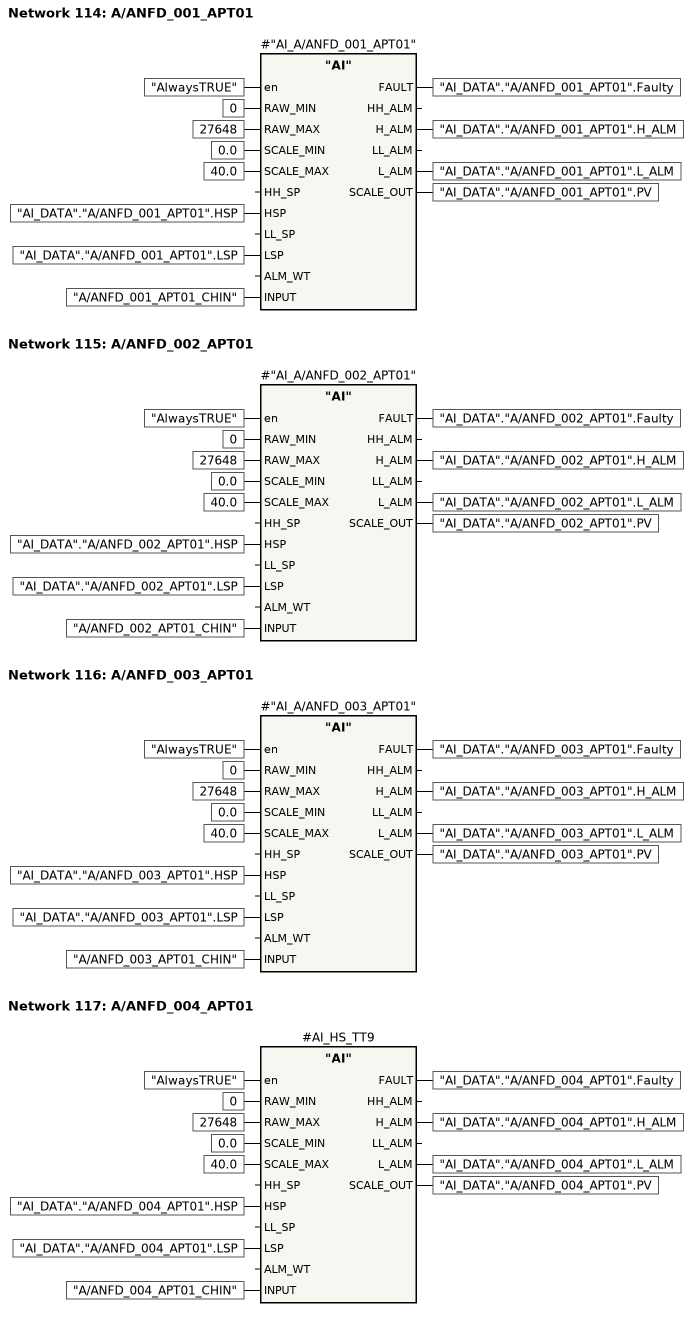
   IF "AlwaysTRUE" THEN
       #"AI_A/ANFD_001_APT01"(RAW_MIN := 0,   // "AI"
                              RAW_MAX := 27648,
                              SCALE_MIN := 0.0,
                              SCALE_MAX := 40.0,
                              HSP := "AI_DATA"."A/ANFD_001_APT01".HSP,
                              LSP := "AI_DATA"."A/ANFD_001_APT01".LSP,
                              INPUT := "A/ANFD_001_APT01_CHIN",
                              FAULT => "AI_DATA"."A/ANFD_001_APT01".Faulty,
                              H_ALM => "AI_DATA"."A/ANFD_001_APT01".H_ALM,
                              L_ALM => "AI_DATA"."A/ANFD_001_APT01".L_ALM,
                              SCALE_OUT => "AI_DATA"."A/ANFD_001_APT01".PV);
   END_IF;
END_REGION

REGION Network 115: A/ANFD_002_APT01
   IF "AlwaysTRUE" THEN
       #"AI_A/ANFD_002_APT01"(RAW_MIN := 0,   // "AI"
                              RAW_MAX := 27648,
                              SCALE_MIN := 0.0,
                              SCALE_MAX := 40.0,
                              HSP := "AI_DATA"."A/ANFD_002_APT01".HSP,
                              LSP := "AI_DATA"."A/ANFD_002_APT01".LSP,
                              INPUT := "A/ANFD_002_APT01_CHIN",
                              FAULT => "AI_DATA"."A/ANFD_002_APT01".Faulty,
                              H_ALM => "AI_DATA"."A/ANFD_002_APT01".H_ALM,
                              L_ALM => "AI_DATA"."A/ANFD_002_APT01".L_ALM,
                              SCALE_OUT => "AI_DATA"."A/ANFD_002_APT01".PV);
   END_IF;
END_REGION

REGION Network 116: A/ANFD_003_APT01
   IF "AlwaysTRUE" THEN
       #"AI_A/ANFD_003_APT01"(RAW_MIN := 0,   // "AI"
                              RAW_MAX := 27648,
                              SCALE_MIN := 0.0,
                              SCALE_MAX := 40.0,
                              HSP := "AI_DATA"."A/ANFD_003_APT01".HSP,
                              LSP := "AI_DATA"."A/ANFD_003_APT01".LSP,
                              INPUT := "A/ANFD_003_APT01_CHIN",
                              FAULT => "AI_DATA"."A/ANFD_003_APT01".Faulty,
                              H_ALM => "AI_DATA"."A/ANFD_003_APT01".H_ALM,
                              L_ALM => "AI_DATA"."A/ANFD_003_APT01".L_ALM,
                              SCALE_OUT => "AI_DATA"."A/ANFD_003_APT01".PV);
   END_IF;
END_REGION

REGION Network 117: A/ANFD_004_APT01
   IF "AlwaysTRUE" THEN
       #AI_HS_TT9(RAW_MIN := 0,   // "AI"
                  RAW_MAX := 27648,
                  SCALE_MIN := 0.0,
                  SCALE_MAX := 40.0,
                  HSP := "AI_DATA"."A/ANFD_004_APT01".HSP,
                  LSP := "AI_DATA"."A/ANFD_004_APT01".LSP,
                  INPUT := "A/ANFD_004_APT01_CHIN",
                  FAULT => "AI_DATA"."A/ANFD_004_APT01".Faulty,
                  H_ALM => "AI_DATA"."A/ANFD_004_APT01".H_ALM,
                  L_ALM => "AI_DATA"."A/ANFD_004_APT01".L_ALM,
                  SCALE_OUT => "AI_DATA"."A/ANFD_004_APT01".PV);
   END_IF;
END_REGION

REGION Network 118: A/ANFD_001_TT01
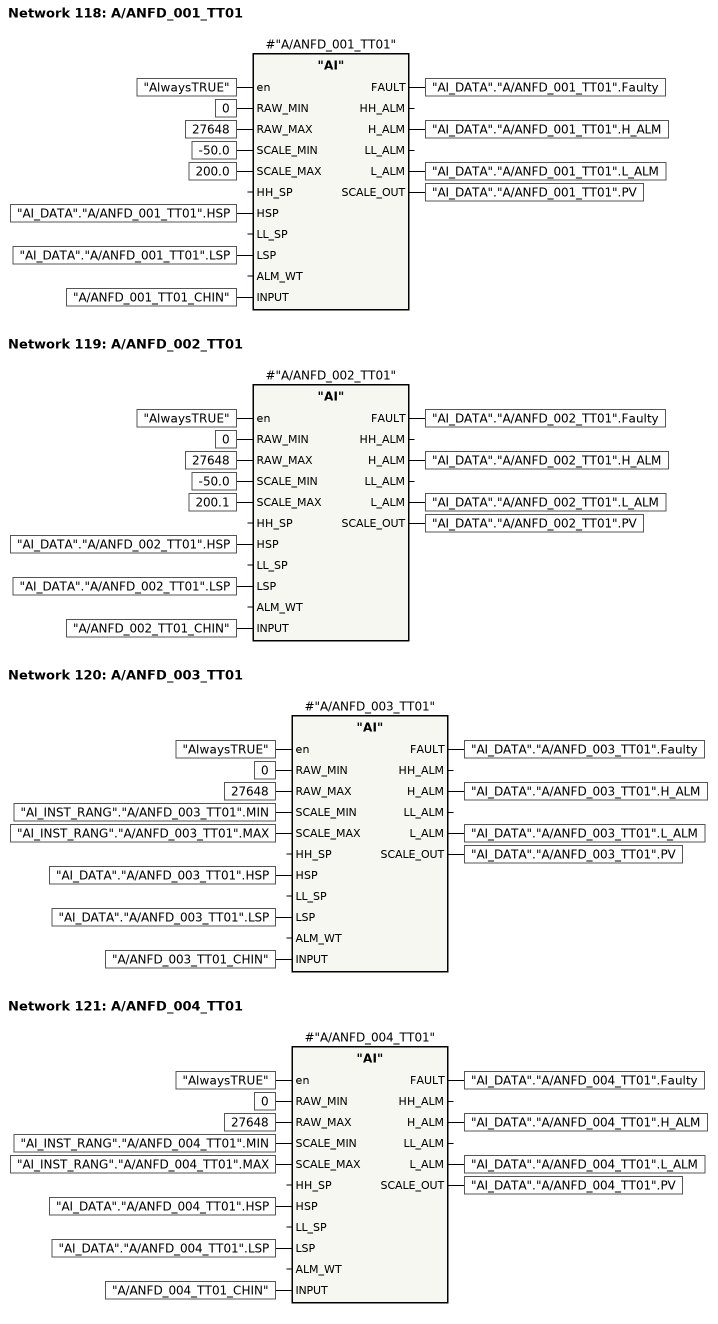
   IF "AlwaysTRUE" THEN
       #"A/ANFD_001_TT01"(RAW_MIN := 0,   // "AI"
                          RAW_MAX := 27648,
                          SCALE_MIN := -50.0,
                          SCALE_MAX := 200.0,
                          HSP := "AI_DATA"."A/ANFD_001_TT01".HSP,
                          LSP := "AI_DATA"."A/ANFD_001_TT01".LSP,
                          INPUT := "A/ANFD_001_TT01_CHIN",
                          FAULT => "AI_DATA"."A/ANFD_001_TT01".Faulty,
                          H_ALM => "AI_DATA"."A/ANFD_001_TT01".H_ALM,
                          L_ALM => "AI_DATA"."A/ANFD_001_TT01".L_ALM,
                          SCALE_OUT => "AI_DATA"."A/ANFD_001_TT01".PV);
   END_IF;
END_REGION

REGION Network 119: A/ANFD_002_TT01
   IF "AlwaysTRUE" THEN
       #"A/ANFD_002_TT01"(RAW_MIN := 0,   // "AI"
                          RAW_MAX := 27648,
                          SCALE_MIN := -50.0,
                          SCALE_MAX := 200.1,
                          HSP := "AI_DATA"."A/ANFD_002_TT01".HSP,
                          LSP := "AI_DATA"."A/ANFD_002_TT01".LSP,
                          INPUT := "A/ANFD_002_TT01_CHIN",
                          FAULT => "AI_DATA"."A/ANFD_002_TT01".Faulty,
                          H_ALM => "AI_DATA"."A/ANFD_002_TT01".H_ALM,
                          L_ALM => "AI_DATA"."A/ANFD_002_TT01".L_ALM,
                          SCALE_OUT => "AI_DATA"."A/ANFD_002_TT01".PV);
   END_IF;
END_REGION

REGION Network 120: A/ANFD_003_TT01
   IF "AlwaysTRUE" THEN
       #"A/ANFD_003_TT01"(RAW_MIN := 0,   // "AI"
                          RAW_MAX := 27648,
                          SCALE_MIN := "AI_INST_RANG"."A/ANFD_003_TT01".MIN,
                          SCALE_MAX := "AI_INST_RANG"."A/ANFD_003_TT01".MAX,
                          HSP := "AI_DATA"."A/ANFD_003_TT01".HSP,
                          LSP := "AI_DATA"."A/ANFD_003_TT01".LSP,
                          INPUT := "A/ANFD_003_TT01_CHIN",
                          FAULT => "AI_DATA"."A/ANFD_003_TT01".Faulty,
                          H_ALM => "AI_DATA"."A/ANFD_003_TT01".H_ALM,
                          L_ALM => "AI_DATA"."A/ANFD_003_TT01".L_ALM,
                          SCALE_OUT => "AI_DATA"."A/ANFD_003_TT01".PV);
   END_IF;
END_REGION

REGION Network 121: A/ANFD_004_TT01
   IF "AlwaysTRUE" THEN
       #"A/ANFD_004_TT01"(RAW_MIN := 0,   // "AI"
                          RAW_MAX := 27648,
                          SCALE_MIN := "AI_INST_RANG"."A/ANFD_004_TT01".MIN,
                          SCALE_MAX := "AI_INST_RANG"."A/ANFD_004_TT01".MAX,
                          HSP := "AI_DATA"."A/ANFD_004_TT01".HSP,
                          LSP := "AI_DATA"."A/ANFD_004_TT01".LSP,
                          INPUT := "A/ANFD_004_TT01_CHIN",
                          FAULT => "AI_DATA"."A/ANFD_004_TT01".Faulty,
                          H_ALM => "AI_DATA"."A/ANFD_004_TT01".H_ALM,
                          L_ALM => "AI_DATA"."A/ANFD_004_TT01".L_ALM,
                          SCALE_OUT => "AI_DATA"."A/ANFD_004_TT01".PV);
   END_IF;
END_REGION

REGION Network 122: RCVD_001_APT01
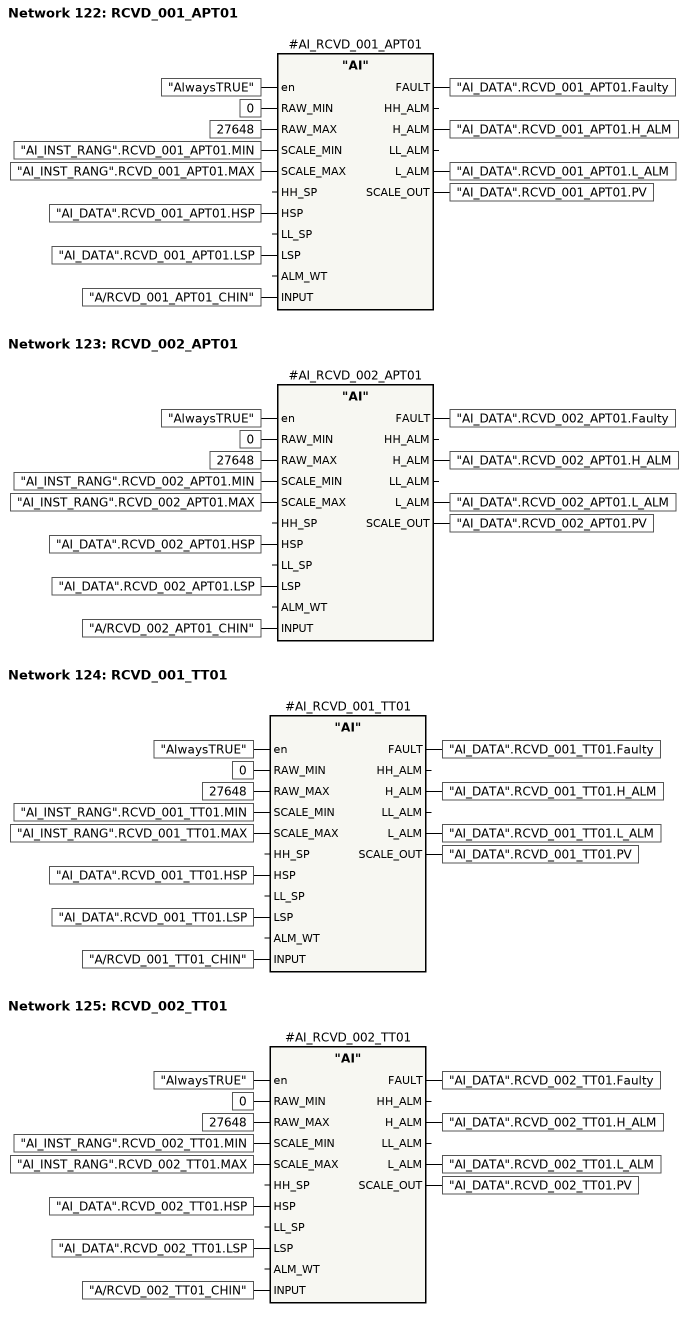
   IF "AlwaysTRUE" THEN
       #AI_RCVD_001_APT01(RAW_MIN := 0,   // "AI"
                          RAW_MAX := 27648,
                          SCALE_MIN := "AI_INST_RANG".RCVD_001_APT01.MIN,
                          SCALE_MAX := "AI_INST_RANG".RCVD_001_APT01.MAX,
                          HSP := "AI_DATA".RCVD_001_APT01.HSP,
                          LSP := "AI_DATA".RCVD_001_APT01.LSP,
                          INPUT := "A/RCVD_001_APT01_CHIN",
                          FAULT => "AI_DATA".RCVD_001_APT01.Faulty,
                          H_ALM => "AI_DATA".RCVD_001_APT01.H_ALM,
                          L_ALM => "AI_DATA".RCVD_001_APT01.L_ALM,
                          SCALE_OUT => "AI_DATA".RCVD_001_APT01.PV);
   END_IF;
END_REGION

REGION Network 123: RCVD_002_APT01
   IF "AlwaysTRUE" THEN
       #AI_RCVD_002_APT01(RAW_MIN := 0,   // "AI"
                          RAW_MAX := 27648,
                          SCALE_MIN := "AI_INST_RANG".RCVD_002_APT01.MIN,
                          SCALE_MAX := "AI_INST_RANG".RCVD_002_APT01.MAX,
                          HSP := "AI_DATA".RCVD_002_APT01.HSP,
                          LSP := "AI_DATA".RCVD_002_APT01.LSP,
                          INPUT := "A/RCVD_002_APT01_CHIN",
                          FAULT => "AI_DATA".RCVD_002_APT01.Faulty,
                          H_ALM => "AI_DATA".RCVD_002_APT01.H_ALM,
                          L_ALM => "AI_DATA".RCVD_002_APT01.L_ALM,
                          SCALE_OUT => "AI_DATA".RCVD_002_APT01.PV);
   END_IF;
END_REGION

REGION Network 124: RCVD_001_TT01
   IF "AlwaysTRUE" THEN
       #AI_RCVD_001_TT01(RAW_MIN := 0,   // "AI"
                         RAW_MAX := 27648,
                         SCALE_MIN := "AI_INST_RANG".RCVD_001_TT01.MIN,
                         SCALE_MAX := "AI_INST_RANG".RCVD_001_TT01.MAX,
                         HSP := "AI_DATA".RCVD_001_TT01.HSP,
                         LSP := "AI_DATA".RCVD_001_TT01.LSP,
                         INPUT := "A/RCVD_001_TT01_CHIN",
                         FAULT => "AI_DATA".RCVD_001_TT01.Faulty,
                         H_ALM => "AI_DATA".RCVD_001_TT01.H_ALM,
                         L_ALM => "AI_DATA".RCVD_001_TT01.L_ALM,
                         SCALE_OUT => "AI_DATA".RCVD_001_TT01.PV);
   END_IF;
END_REGION

REGION Network 125: RCVD_002_TT01
   IF "AlwaysTRUE" THEN
       #AI_RCVD_002_TT01(RAW_MIN := 0,   // "AI"
                         RAW_MAX := 27648,
                         SCALE_MIN := "AI_INST_RANG".RCVD_002_TT01.MIN,
                         SCALE_MAX := "AI_INST_RANG".RCVD_002_TT01.MAX,
                         HSP := "AI_DATA".RCVD_002_TT01.HSP,
                         LSP := "AI_DATA".RCVD_002_TT01.LSP,
                         INPUT := "A/RCVD_002_TT01_CHIN",
                         FAULT => "AI_DATA".RCVD_002_TT01.Faulty,
                         H_ALM => "AI_DATA".RCVD_002_TT01.H_ALM,
                         L_ALM => "AI_DATA".RCVD_002_TT01.L_ALM,
                         SCALE_OUT => "AI_DATA".RCVD_002_TT01.PV);
   END_IF;
END_REGION

REGION Network 126: A/VTD_001_APT01
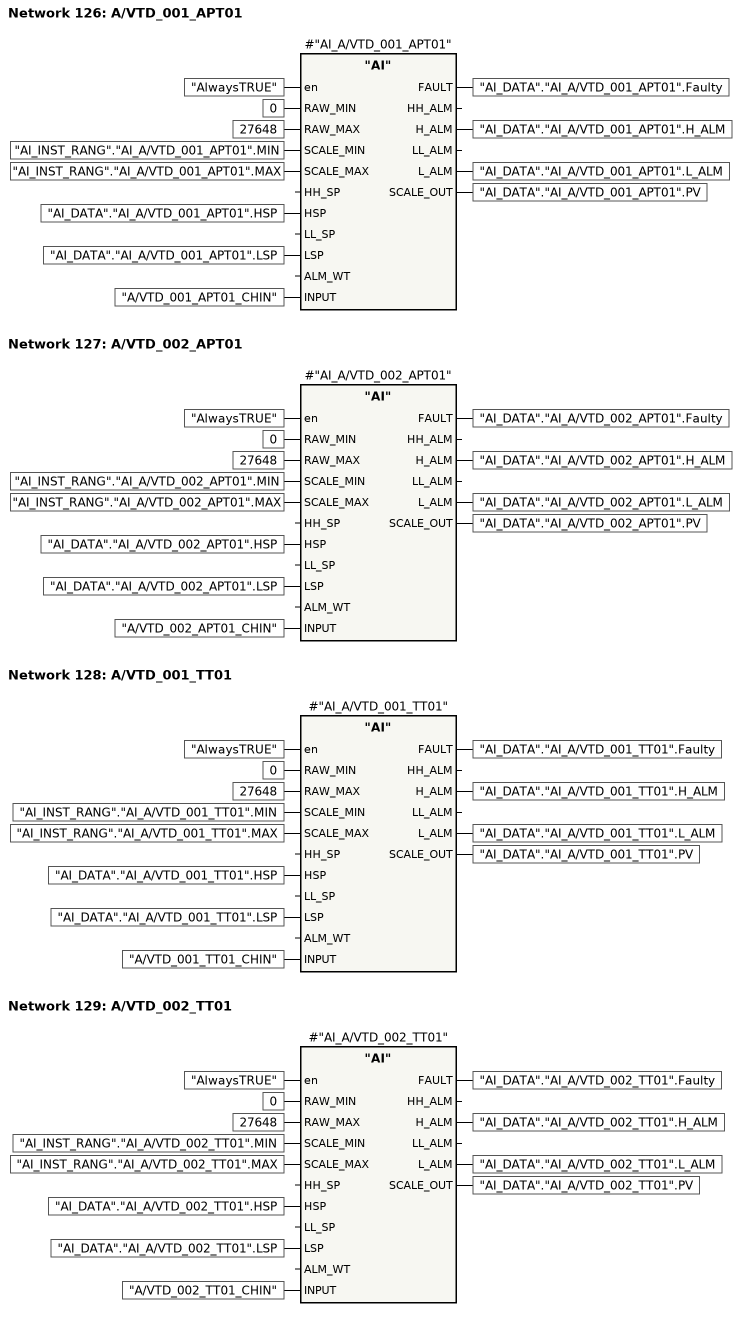
   IF "AlwaysTRUE" THEN
       #"AI_A/VTD_001_APT01"(RAW_MIN := 0,   // "AI"
                             RAW_MAX := 27648,
                             SCALE_MIN := "AI_INST_RANG"."AI_A/VTD_001_APT01".MIN,
                             SCALE_MAX := "AI_INST_RANG"."AI_A/VTD_001_APT01".MAX,
                             HSP := "AI_DATA"."AI_A/VTD_001_APT01".HSP,
                             LSP := "AI_DATA"."AI_A/VTD_001_APT01".LSP,
                             INPUT := "A/VTD_001_APT01_CHIN",
                             FAULT => "AI_DATA"."AI_A/VTD_001_APT01".Faulty,
                             H_ALM => "AI_DATA"."AI_A/VTD_001_APT01".H_ALM,
                             L_ALM => "AI_DATA"."AI_A/VTD_001_APT01".L_ALM,
                             SCALE_OUT => "AI_DATA"."AI_A/VTD_001_APT01".PV);
   END_IF;
END_REGION

REGION Network 127: A/VTD_002_APT01
   IF "AlwaysTRUE" THEN
       #"AI_A/VTD_002_APT01"(RAW_MIN := 0,   // "AI"
                             RAW_MAX := 27648,
                             SCALE_MIN := "AI_INST_RANG"."AI_A/VTD_002_APT01".MIN,
                             SCALE_MAX := "AI_INST_RANG"."AI_A/VTD_002_APT01".MAX,
                             HSP := "AI_DATA"."AI_A/VTD_002_APT01".HSP,
                             LSP := "AI_DATA"."AI_A/VTD_002_APT01".LSP,
                             INPUT := "A/VTD_002_APT01_CHIN",
                             FAULT => "AI_DATA"."AI_A/VTD_002_APT01".Faulty,
                             H_ALM => "AI_DATA"."AI_A/VTD_002_APT01".H_ALM,
                             L_ALM => "AI_DATA"."AI_A/VTD_002_APT01".L_ALM,
                             SCALE_OUT => "AI_DATA"."AI_A/VTD_002_APT01".PV);
   END_IF;
END_REGION

REGION Network 128: A/VTD_001_TT01
   IF "AlwaysTRUE" THEN
       #"AI_A/VTD_001_TT01"(RAW_MIN := 0,   // "AI"
                            RAW_MAX := 27648,
                            SCALE_MIN := "AI_INST_RANG"."AI_A/VTD_001_TT01".MIN,
                            SCALE_MAX := "AI_INST_RANG"."AI_A/VTD_001_TT01".MAX,
                            HSP := "AI_DATA"."AI_A/VTD_001_TT01".HSP,
                            LSP := "AI_DATA"."AI_A/VTD_001_TT01".LSP,
                            INPUT := "A/VTD_001_TT01_CHIN",
                            FAULT => "AI_DATA"."AI_A/VTD_001_TT01".Faulty,
                            H_ALM => "AI_DATA"."AI_A/VTD_001_TT01".H_ALM,
                            L_ALM => "AI_DATA"."AI_A/VTD_001_TT01".L_ALM,
                            SCALE_OUT => "AI_DATA"."AI_A/VTD_001_TT01".PV);
   END_IF;
END_REGION

REGION Network 129: A/VTD_002_TT01
   IF "AlwaysTRUE" THEN
       #"AI_A/VTD_002_TT01"(RAW_MIN := 0,   // "AI"
                            RAW_MAX := 27648,
                            SCALE_MIN := "AI_INST_RANG"."AI_A/VTD_002_TT01".MIN,
                            SCALE_MAX := "AI_INST_RANG"."AI_A/VTD_002_TT01".MAX,
                            HSP := "AI_DATA"."AI_A/VTD_002_TT01".HSP,
                            LSP := "AI_DATA"."AI_A/VTD_002_TT01".LSP,
                            INPUT := "A/VTD_002_TT01_CHIN",
                            FAULT => "AI_DATA"."AI_A/VTD_002_TT01".Faulty,
                            H_ALM => "AI_DATA"."AI_A/VTD_002_TT01".H_ALM,
                            L_ALM => "AI_DATA"."AI_A/VTD_002_TT01".L_ALM,
                            SCALE_OUT => "AI_DATA"."AI_A/VTD_002_TT01".PV);
   END_IF;
END_REGION

REGION Network 130: A/TD_001_TT01
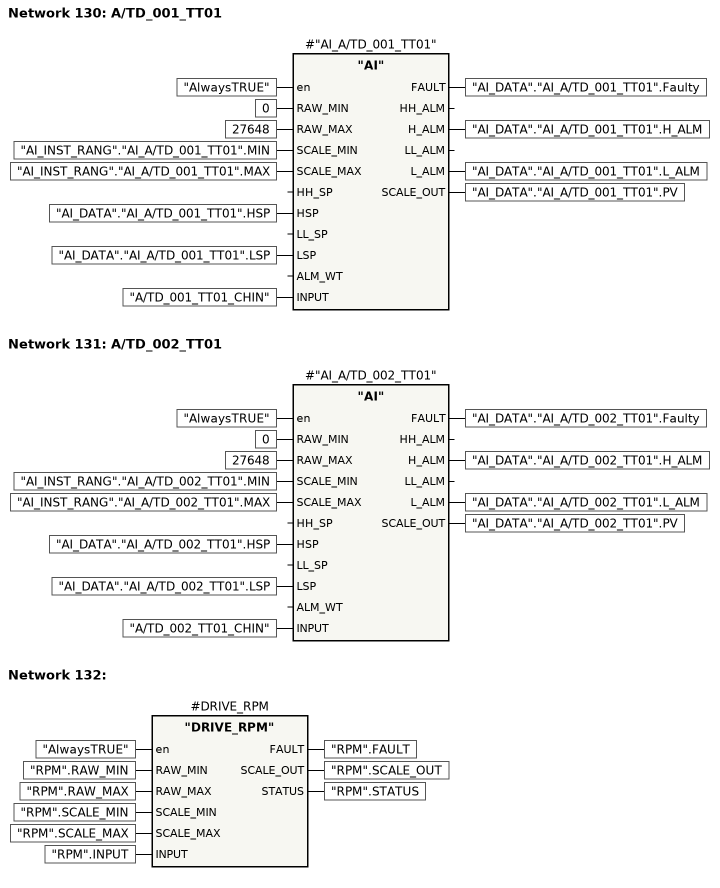
   IF "AlwaysTRUE" THEN
       #"AI_A/TD_001_TT01"(RAW_MIN := 0,   // "AI"
                           RAW_MAX := 27648,
                           SCALE_MIN := "AI_INST_RANG"."AI_A/TD_001_TT01".MIN,
                           SCALE_MAX := "AI_INST_RANG"."AI_A/TD_001_TT01".MAX,
                           HSP := "AI_DATA"."AI_A/TD_001_TT01".HSP,
                           LSP := "AI_DATA"."AI_A/TD_001_TT01".LSP,
                           INPUT := "A/TD_001_TT01_CHIN",
                           FAULT => "AI_DATA"."AI_A/TD_001_TT01".Faulty,
                           H_ALM => "AI_DATA"."AI_A/TD_001_TT01".H_ALM,
                           L_ALM => "AI_DATA"."AI_A/TD_001_TT01".L_ALM,
                           SCALE_OUT => "AI_DATA"."AI_A/TD_001_TT01".PV);
   END_IF;
END_REGION

REGION Network 131: A/TD_002_TT01
   IF "AlwaysTRUE" THEN
       #"AI_A/TD_002_TT01"(RAW_MIN := 0,   // "AI"
                           RAW_MAX := 27648,
                           SCALE_MIN := "AI_INST_RANG"."AI_A/TD_002_TT01".MIN,
                           SCALE_MAX := "AI_INST_RANG"."AI_A/TD_002_TT01".MAX,
                           HSP := "AI_DATA"."AI_A/TD_002_TT01".HSP,
                           LSP := "AI_DATA"."AI_A/TD_002_TT01".LSP,
                           INPUT := "A/TD_002_TT01_CHIN",
                           FAULT => "AI_DATA"."AI_A/TD_002_TT01".Faulty,
                           H_ALM => "AI_DATA"."AI_A/TD_002_TT01".H_ALM,
                           L_ALM => "AI_DATA"."AI_A/TD_002_TT01".L_ALM,
                           SCALE_OUT => "AI_DATA"."AI_A/TD_002_TT01".PV);
   END_IF;
END_REGION

REGION Network 132
   IF "AlwaysTRUE" THEN
       #DRIVE_RPM(RAW_MIN := "RPM".RAW_MIN,   // "DRIVE_RPM"
                  RAW_MAX := "RPM".RAW_MAX,
                  SCALE_MIN := "RPM".SCALE_MIN,
                  SCALE_MAX := "RPM".SCALE_MAX,
                  INPUT := "RPM".INPUT,
                  FAULT => "RPM".FAULT,
                  SCALE_OUT => "RPM".SCALE_OUT,
                  STATUS => "RPM".STATUS);
   END_IF;
END_REGION

REGION Network 133 (SCL)
   "RPM".INPUT[1] := "GLR_001";
   "RPM".INPUT[2] := "SSR_002";
   "RPM".INPUT[3] := "SSR_003";
   "RPM".INPUT[4] := "SSR_004";
   "RPM".INPUT[5] := "GLR_005";
   "RPM".INPUT[6] := "GLR_006";
   "RPM".INPUT[7] := "SSR_007";
   "RPM".INPUT[8] := "SSR_008";
   "RPM".INPUT[9] := "GLR_009";
   "RPM".INPUT[10] := "GLR_010";
   "RPM".INPUT[11] := "SSR_011";
   "RPM".INPUT[12] := "GLR_012";
   "RPM".INPUT[13] := "SSR_013";
   "RPM".INPUT[14] := "SSR_014";
   "RPM".INPUT[15] := "SSR_015";
   "RPM".INPUT[16] := "GLR_016";
   "RPM".INPUT[17] := "SSR_017";
   "RPM".INPUT[18] := "GLR_018";
END_REGION
END_FUNCTION_BLOCK
